(* IEC 61131-3 sources: sis-interlock-demo/tests/POUs/Generated/FB_VoteTruth_Test (part 2) *)

(* ---- Fb2oo2DADIMatchesTable.method.impl.st ---- *)
// AUTO-GENERATED by cemgen 1.0.0 — не редактировать: правьте матрицу и запустите
//   python -m cemgen generate <файл матрицы .csv или .xlsx>
// Матрица: SIS-V101-CEM, объект V-101, ревизия B от 2026-10-19, SHA-256 сетки df2ed4841a9453ca
coUnit.TEST('VoteTruth_Fb2oo2DADI_MatchesTable');
stCfg.eArch := E_VoteArch.Vote2oo2;
stCfg.ePolicy := E_DegradePolicy.DegradeAvailable;
stCfg.eInput := E_SisInputKind.Discrete;
stCfg.xDiHealthy := TRUE;
stCfg.eLimitDir := E_LimitDir.High;
stCfg.rTripLimit_eu := 50.0;
stCfg.rHyst_eu := 0.0;
stCfg.rDiscrepancyMax_eu := 0.0;
stCfg.tDiscrepancyDelay := T#0S;
stCfg.tBypassMax := T#1H;
stCfg.uiMaxBypass := 1;
FOR uiRow := 0 TO 63 DO
    RowInputs(uiRow := uiRow, uiChannels := 2, xBypass := FALSE, stIn := stIn, stCmd := stCmd);
    fbVote(stIn := stIn, stCmd := stCmd, stCfg := stCfg, xBypassPermit := TRUE, uiCause := 1,
        itfTime := fbTime);
    RowInputs(uiRow := uiRow, uiChannels := 2, xBypass := TRUE, stIn := stIn, stCmd := stCmd);
    fbVote(stIn := stIn, stCmd := stCmd, stCfg := stCfg, xBypassPermit := TRUE, uiCause := 1,
        itfTime := fbTime);
    bAct := EncodeFb(xTrip := fbVote.xTrip, stSts := fbVote.stSts);
    bExp := GVL_VoteTruthTable.TT_FB_2OO2_DA_DI[uiRow];
    xMiss := bAct <> bExp;
    xFirst := xMiss AND uiMismatch = 0;
    uiFirstRow := SEL(xFirst, uiFirstRow, uiRow);
    bFirstExp := SEL(xFirst, bFirstExp, bExp);
    bFirstAct := SEL(xFirst, bFirstAct, bAct);
    uiMismatch := uiMismatch + BOOL_TO_UINT(xMiss);
END_FOR
AssertEquals_UINT(Expected := 0, Actual := uiMismatch,
    Message := MismatchText(sTable := 'TT_FB_2OO2_DA_DI', uiRow := uiFirstRow, bExpected := bFirstExp,
        bActual := bFirstAct));
coUnit.TEST_FINISHED();

(* ---- Fb2oo2DSAIMatchesTable.method.decl.st ---- *)
// AUTO-GENERATED by cemgen 1.0.0 — не редактировать: правьте матрицу и запустите
//   python -m cemgen generate <файл матрицы .csv или .xlsx>
// Матрица: SIS-V101-CEM, объект V-101, ревизия B от 2026-10-19, SHA-256 сетки df2ed4841a9453ca
// Назначение: тест VoteTruth_Fb2oo2DSAI_MatchesTable набора FB_VoteTruth_Test.
// Автор:      kr0nsch; код — генератор cemgen
// Версия:     1.0.0
// Документ:   docs/DESIGN.md, раздел «10. Генератор cemgen»; docs/cause_effect_matrix.md
// ВНИМАНИЕ:   код демонстрационный и не предназначен для систем безопасности. Реальная ПАЗ требует
//             определения SIL, сертифицированных аппаратных и программных средств и валидации по
//             ГОСТ Р МЭК 61511.
// FB_Voting, схема 2oo2, политика DegradeSafe, аналоговые каналы: все 64 сочетаний «требование ×
// достоверность × запрос байпаса» совпадают с таблицей TT_FB_2OO2_DS_AI. На строку — два вызова одного
// экземпляра: без запросов байпаса (сброс байпасов прошлой строки) и с полной строкой.
METHOD PRIVATE Fb2oo2DSAIMatchesTable
VAR
    fbTime     : PL.FB_FakeTime;   // время не меняется
    fbVote     : FB_Voting;        // ФБ под тестом, один экземпляр на все строки
    stCfg      : ST_VotingCfg;     // конфигурация теста уровня 2
    stIn       : ST_VoteIn;        // входы строки
    stCmd      : ST_VoteCmd;       // запросы байпаса строки
    uiRow      : UINT;             // строка таблицы
    bAct       : BYTE;             // фактический байт результата
    bExp       : BYTE;             // ожидаемый байт из таблицы
    xMiss      : BOOL;             // строка не совпала
    xFirst     : BOOL;             // первая несовпавшая строка
    uiMismatch : UINT;             // несовпавших строк
    uiFirstRow : UINT;             // первая несовпавшая строка
    bFirstExp  : BYTE;             // ожидаемый байт первой несовпавшей строки
    bFirstAct  : BYTE;             // фактический байт первой несовпавшей строки
END_VAR

(* ---- Fb2oo2DSAIMatchesTable.method.impl.st ---- *)
// AUTO-GENERATED by cemgen 1.0.0 — не редактировать: правьте матрицу и запустите
//   python -m cemgen generate <файл матрицы .csv или .xlsx>
// Матрица: SIS-V101-CEM, объект V-101, ревизия B от 2026-10-19, SHA-256 сетки df2ed4841a9453ca
coUnit.TEST('VoteTruth_Fb2oo2DSAI_MatchesTable');
stCfg.eArch := E_VoteArch.Vote2oo2;
stCfg.ePolicy := E_DegradePolicy.DegradeSafe;
stCfg.eInput := E_SisInputKind.Analog;
stCfg.xDiHealthy := TRUE;
stCfg.eLimitDir := E_LimitDir.High;
stCfg.rTripLimit_eu := 50.0;
stCfg.rHyst_eu := 0.0;
stCfg.rDiscrepancyMax_eu := 0.0;
stCfg.tDiscrepancyDelay := T#0S;
stCfg.tBypassMax := T#1H;
stCfg.uiMaxBypass := 1;
FOR uiRow := 0 TO 63 DO
    RowInputs(uiRow := uiRow, uiChannels := 2, xBypass := FALSE, stIn := stIn, stCmd := stCmd);
    fbVote(stIn := stIn, stCmd := stCmd, stCfg := stCfg, xBypassPermit := TRUE, uiCause := 1,
        itfTime := fbTime);
    RowInputs(uiRow := uiRow, uiChannels := 2, xBypass := TRUE, stIn := stIn, stCmd := stCmd);
    fbVote(stIn := stIn, stCmd := stCmd, stCfg := stCfg, xBypassPermit := TRUE, uiCause := 1,
        itfTime := fbTime);
    bAct := EncodeFb(xTrip := fbVote.xTrip, stSts := fbVote.stSts);
    bExp := GVL_VoteTruthTable.TT_FB_2OO2_DS_AI[uiRow];
    xMiss := bAct <> bExp;
    xFirst := xMiss AND uiMismatch = 0;
    uiFirstRow := SEL(xFirst, uiFirstRow, uiRow);
    bFirstExp := SEL(xFirst, bFirstExp, bExp);
    bFirstAct := SEL(xFirst, bFirstAct, bAct);
    uiMismatch := uiMismatch + BOOL_TO_UINT(xMiss);
END_FOR
AssertEquals_UINT(Expected := 0, Actual := uiMismatch,
    Message := MismatchText(sTable := 'TT_FB_2OO2_DS_AI', uiRow := uiFirstRow, bExpected := bFirstExp,
        bActual := bFirstAct));
coUnit.TEST_FINISHED();

(* ---- Fb2oo2DSDIMatchesTable.method.decl.st ---- *)
// AUTO-GENERATED by cemgen 1.0.0 — не редактировать: правьте матрицу и запустите
//   python -m cemgen generate <файл матрицы .csv или .xlsx>
// Матрица: SIS-V101-CEM, объект V-101, ревизия B от 2026-10-19, SHA-256 сетки df2ed4841a9453ca
// Назначение: тест VoteTruth_Fb2oo2DSDI_MatchesTable набора FB_VoteTruth_Test.
// Автор:      kr0nsch; код — генератор cemgen
// Версия:     1.0.0
// Документ:   docs/DESIGN.md, раздел «10. Генератор cemgen»; docs/cause_effect_matrix.md
// ВНИМАНИЕ:   код демонстрационный и не предназначен для систем безопасности. Реальная ПАЗ требует
//             определения SIL, сертифицированных аппаратных и программных средств и валидации по
//             ГОСТ Р МЭК 61511.
// FB_Voting, схема 2oo2, политика DegradeSafe, дискретные каналы: все 64 сочетаний «требование ×
// достоверность × запрос байпаса» совпадают с таблицей TT_FB_2OO2_DS_DI. На строку — два вызова одного
// экземпляра: без запросов байпаса (сброс байпасов прошлой строки) и с полной строкой.
METHOD PRIVATE Fb2oo2DSDIMatchesTable
VAR
    fbTime     : PL.FB_FakeTime;   // время не меняется
    fbVote     : FB_Voting;        // ФБ под тестом, один экземпляр на все строки
    stCfg      : ST_VotingCfg;     // конфигурация теста уровня 2
    stIn       : ST_VoteIn;        // входы строки
    stCmd      : ST_VoteCmd;       // запросы байпаса строки
    uiRow      : UINT;             // строка таблицы
    bAct       : BYTE;             // фактический байт результата
    bExp       : BYTE;             // ожидаемый байт из таблицы
    xMiss      : BOOL;             // строка не совпала
    xFirst     : BOOL;             // первая несовпавшая строка
    uiMismatch : UINT;             // несовпавших строк
    uiFirstRow : UINT;             // первая несовпавшая строка
    bFirstExp  : BYTE;             // ожидаемый байт первой несовпавшей строки
    bFirstAct  : BYTE;             // фактический байт первой несовпавшей строки
END_VAR

(* ---- Fb2oo2DSDIMatchesTable.method.impl.st ---- *)
// AUTO-GENERATED by cemgen 1.0.0 — не редактировать: правьте матрицу и запустите
//   python -m cemgen generate <файл матрицы .csv или .xlsx>
// Матрица: SIS-V101-CEM, объект V-101, ревизия B от 2026-10-19, SHA-256 сетки df2ed4841a9453ca
coUnit.TEST('VoteTruth_Fb2oo2DSDI_MatchesTable');
stCfg.eArch := E_VoteArch.Vote2oo2;
stCfg.ePolicy := E_DegradePolicy.DegradeSafe;
stCfg.eInput := E_SisInputKind.Discrete;
stCfg.xDiHealthy := TRUE;
stCfg.eLimitDir := E_LimitDir.High;
stCfg.rTripLimit_eu := 50.0;
stCfg.rHyst_eu := 0.0;
stCfg.rDiscrepancyMax_eu := 0.0;
stCfg.tDiscrepancyDelay := T#0S;
stCfg.tBypassMax := T#1H;
stCfg.uiMaxBypass := 1;
FOR uiRow := 0 TO 63 DO
    RowInputs(uiRow := uiRow, uiChannels := 2, xBypass := FALSE, stIn := stIn, stCmd := stCmd);
    fbVote(stIn := stIn, stCmd := stCmd, stCfg := stCfg, xBypassPermit := TRUE, uiCause := 1,
        itfTime := fbTime);
    RowInputs(uiRow := uiRow, uiChannels := 2, xBypass := TRUE, stIn := stIn, stCmd := stCmd);
    fbVote(stIn := stIn, stCmd := stCmd, stCfg := stCfg, xBypassPermit := TRUE, uiCause := 1,
        itfTime := fbTime);
    bAct := EncodeFb(xTrip := fbVote.xTrip, stSts := fbVote.stSts);
    bExp := GVL_VoteTruthTable.TT_FB_2OO2_DS_DI[uiRow];
    xMiss := bAct <> bExp;
    xFirst := xMiss AND uiMismatch = 0;
    uiFirstRow := SEL(xFirst, uiFirstRow, uiRow);
    bFirstExp := SEL(xFirst, bFirstExp, bExp);
    bFirstAct := SEL(xFirst, bFirstAct, bAct);
    uiMismatch := uiMismatch + BOOL_TO_UINT(xMiss);
END_FOR
AssertEquals_UINT(Expected := 0, Actual := uiMismatch,
    Message := MismatchText(sTable := 'TT_FB_2OO2_DS_DI', uiRow := uiFirstRow, bExpected := bFirstExp,
        bActual := bFirstAct));
coUnit.TEST_FINISHED();

(* ---- Fb2oo2VTAIMatchesTable.method.decl.st ---- *)
// AUTO-GENERATED by cemgen 1.0.0 — не редактировать: правьте матрицу и запустите
//   python -m cemgen generate <файл матрицы .csv или .xlsx>
// Матрица: SIS-V101-CEM, объект V-101, ревизия B от 2026-10-19, SHA-256 сетки df2ed4841a9453ca
// Назначение: тест VoteTruth_Fb2oo2VTAI_MatchesTable набора FB_VoteTruth_Test.
// Автор:      kr0nsch; код — генератор cemgen
// Версия:     1.0.0
// Документ:   docs/DESIGN.md, раздел «10. Генератор cemgen»; docs/cause_effect_matrix.md
// ВНИМАНИЕ:   код демонстрационный и не предназначен для систем безопасности. Реальная ПАЗ требует
//             определения SIL, сертифицированных аппаратных и программных средств и валидации по
//             ГОСТ Р МЭК 61511.
// FB_Voting, схема 2oo2, политика VoteTrip, аналоговые каналы: все 64 сочетаний «требование ×
// достоверность × запрос байпаса» совпадают с таблицей TT_FB_2OO2_VT_AI. На строку — два вызова одного
// экземпляра: без запросов байпаса (сброс байпасов прошлой строки) и с полной строкой.
METHOD PRIVATE Fb2oo2VTAIMatchesTable
VAR
    fbTime     : PL.FB_FakeTime;   // время не меняется
    fbVote     : FB_Voting;        // ФБ под тестом, один экземпляр на все строки
    stCfg      : ST_VotingCfg;     // конфигурация теста уровня 2
    stIn       : ST_VoteIn;        // входы строки
    stCmd      : ST_VoteCmd;       // запросы байпаса строки
    uiRow      : UINT;             // строка таблицы
    bAct       : BYTE;             // фактический байт результата
    bExp       : BYTE;             // ожидаемый байт из таблицы
    xMiss      : BOOL;             // строка не совпала
    xFirst     : BOOL;             // первая несовпавшая строка
    uiMismatch : UINT;             // несовпавших строк
    uiFirstRow : UINT;             // первая несовпавшая строка
    bFirstExp  : BYTE;             // ожидаемый байт первой несовпавшей строки
    bFirstAct  : BYTE;             // фактический байт первой несовпавшей строки
END_VAR

(* ---- Fb2oo2VTAIMatchesTable.method.impl.st ---- *)
// AUTO-GENERATED by cemgen 1.0.0 — не редактировать: правьте матрицу и запустите
//   python -m cemgen generate <файл матрицы .csv или .xlsx>
// Матрица: SIS-V101-CEM, объект V-101, ревизия B от 2026-10-19, SHA-256 сетки df2ed4841a9453ca
coUnit.TEST('VoteTruth_Fb2oo2VTAI_MatchesTable');
stCfg.eArch := E_VoteArch.Vote2oo2;
stCfg.ePolicy := E_DegradePolicy.VoteTrip;
stCfg.eInput := E_SisInputKind.Analog;
stCfg.xDiHealthy := TRUE;
stCfg.eLimitDir := E_LimitDir.High;
stCfg.rTripLimit_eu := 50.0;
stCfg.rHyst_eu := 0.0;
stCfg.rDiscrepancyMax_eu := 0.0;
stCfg.tDiscrepancyDelay := T#0S;
stCfg.tBypassMax := T#1H;
stCfg.uiMaxBypass := 1;
FOR uiRow := 0 TO 63 DO
    RowInputs(uiRow := uiRow, uiChannels := 2, xBypass := FALSE, stIn := stIn, stCmd := stCmd);
    fbVote(stIn := stIn, stCmd := stCmd, stCfg := stCfg, xBypassPermit := TRUE, uiCause := 1,
        itfTime := fbTime);
    RowInputs(uiRow := uiRow, uiChannels := 2, xBypass := TRUE, stIn := stIn, stCmd := stCmd);
    fbVote(stIn := stIn, stCmd := stCmd, stCfg := stCfg, xBypassPermit := TRUE, uiCause := 1,
        itfTime := fbTime);
    bAct := EncodeFb(xTrip := fbVote.xTrip, stSts := fbVote.stSts);
    bExp := GVL_VoteTruthTable.TT_FB_2OO2_VT_AI[uiRow];
    xMiss := bAct <> bExp;
    xFirst := xMiss AND uiMismatch = 0;
    uiFirstRow := SEL(xFirst, uiFirstRow, uiRow);
    bFirstExp := SEL(xFirst, bFirstExp, bExp);
    bFirstAct := SEL(xFirst, bFirstAct, bAct);
    uiMismatch := uiMismatch + BOOL_TO_UINT(xMiss);
END_FOR
AssertEquals_UINT(Expected := 0, Actual := uiMismatch,
    Message := MismatchText(sTable := 'TT_FB_2OO2_VT_AI', uiRow := uiFirstRow, bExpected := bFirstExp,
        bActual := bFirstAct));
coUnit.TEST_FINISHED();

(* ---- Fb2oo2VTDIMatchesTable.method.decl.st ---- *)
// AUTO-GENERATED by cemgen 1.0.0 — не редактировать: правьте матрицу и запустите
//   python -m cemgen generate <файл матрицы .csv или .xlsx>
// Матрица: SIS-V101-CEM, объект V-101, ревизия B от 2026-10-19, SHA-256 сетки df2ed4841a9453ca
// Назначение: тест VoteTruth_Fb2oo2VTDI_MatchesTable набора FB_VoteTruth_Test.
// Автор:      kr0nsch; код — генератор cemgen
// Версия:     1.0.0
// Документ:   docs/DESIGN.md, раздел «10. Генератор cemgen»; docs/cause_effect_matrix.md
// ВНИМАНИЕ:   код демонстрационный и не предназначен для систем безопасности. Реальная ПАЗ требует
//             определения SIL, сертифицированных аппаратных и программных средств и валидации по
//             ГОСТ Р МЭК 61511.
// FB_Voting, схема 2oo2, политика VoteTrip, дискретные каналы: все 64 сочетаний «требование ×
// достоверность × запрос байпаса» совпадают с таблицей TT_FB_2OO2_VT_DI. На строку — два вызова одного
// экземпляра: без запросов байпаса (сброс байпасов прошлой строки) и с полной строкой.
METHOD PRIVATE Fb2oo2VTDIMatchesTable
VAR
    fbTime     : PL.FB_FakeTime;   // время не меняется
    fbVote     : FB_Voting;        // ФБ под тестом, один экземпляр на все строки
    stCfg      : ST_VotingCfg;     // конфигурация теста уровня 2
    stIn       : ST_VoteIn;        // входы строки
    stCmd      : ST_VoteCmd;       // запросы байпаса строки
    uiRow      : UINT;             // строка таблицы
    bAct       : BYTE;             // фактический байт результата
    bExp       : BYTE;             // ожидаемый байт из таблицы
    xMiss      : BOOL;             // строка не совпала
    xFirst     : BOOL;             // первая несовпавшая строка
    uiMismatch : UINT;             // несовпавших строк
    uiFirstRow : UINT;             // первая несовпавшая строка
    bFirstExp  : BYTE;             // ожидаемый байт первой несовпавшей строки
    bFirstAct  : BYTE;             // фактический байт первой несовпавшей строки
END_VAR

(* ---- Fb2oo2VTDIMatchesTable.method.impl.st ---- *)
// AUTO-GENERATED by cemgen 1.0.0 — не редактировать: правьте матрицу и запустите
//   python -m cemgen generate <файл матрицы .csv или .xlsx>
// Матрица: SIS-V101-CEM, объект V-101, ревизия B от 2026-10-19, SHA-256 сетки df2ed4841a9453ca
coUnit.TEST('VoteTruth_Fb2oo2VTDI_MatchesTable');
stCfg.eArch := E_VoteArch.Vote2oo2;
stCfg.ePolicy := E_DegradePolicy.VoteTrip;
stCfg.eInput := E_SisInputKind.Discrete;
stCfg.xDiHealthy := TRUE;
stCfg.eLimitDir := E_LimitDir.High;
stCfg.rTripLimit_eu := 50.0;
stCfg.rHyst_eu := 0.0;
stCfg.rDiscrepancyMax_eu := 0.0;
stCfg.tDiscrepancyDelay := T#0S;
stCfg.tBypassMax := T#1H;
stCfg.uiMaxBypass := 1;
FOR uiRow := 0 TO 63 DO
    RowInputs(uiRow := uiRow, uiChannels := 2, xBypass := FALSE, stIn := stIn, stCmd := stCmd);
    fbVote(stIn := stIn, stCmd := stCmd, stCfg := stCfg, xBypassPermit := TRUE, uiCause := 1,
        itfTime := fbTime);
    RowInputs(uiRow := uiRow, uiChannels := 2, xBypass := TRUE, stIn := stIn, stCmd := stCmd);
    fbVote(stIn := stIn, stCmd := stCmd, stCfg := stCfg, xBypassPermit := TRUE, uiCause := 1,
        itfTime := fbTime);
    bAct := EncodeFb(xTrip := fbVote.xTrip, stSts := fbVote.stSts);
    bExp := GVL_VoteTruthTable.TT_FB_2OO2_VT_DI[uiRow];
    xMiss := bAct <> bExp;
    xFirst := xMiss AND uiMismatch = 0;
    uiFirstRow := SEL(xFirst, uiFirstRow, uiRow);
    bFirstExp := SEL(xFirst, bFirstExp, bExp);
    bFirstAct := SEL(xFirst, bFirstAct, bAct);
    uiMismatch := uiMismatch + BOOL_TO_UINT(xMiss);
END_FOR
AssertEquals_UINT(Expected := 0, Actual := uiMismatch,
    Message := MismatchText(sTable := 'TT_FB_2OO2_VT_DI', uiRow := uiFirstRow, bExpected := bFirstExp,
        bActual := bFirstAct));
coUnit.TEST_FINISHED();

(* ---- Fb2oo3DAAIMatchesTable.method.decl.st ---- *)
// AUTO-GENERATED by cemgen 1.0.0 — не редактировать: правьте матрицу и запустите
//   python -m cemgen generate <файл матрицы .csv или .xlsx>
// Матрица: SIS-V101-CEM, объект V-101, ревизия B от 2026-10-19, SHA-256 сетки df2ed4841a9453ca
// Назначение: тест VoteTruth_Fb2oo3DAAI_MatchesTable набора FB_VoteTruth_Test.
// Автор:      kr0nsch; код — генератор cemgen
// Версия:     1.0.0
// Документ:   docs/DESIGN.md, раздел «10. Генератор cemgen»; docs/cause_effect_matrix.md
// ВНИМАНИЕ:   код демонстрационный и не предназначен для систем безопасности. Реальная ПАЗ требует
//             определения SIL, сертифицированных аппаратных и программных средств и валидации по
//             ГОСТ Р МЭК 61511.
// FB_Voting, схема 2oo3, политика DegradeAvailable, аналоговые каналы: все 512 сочетаний «требование ×
// достоверность × запрос байпаса» совпадают с таблицей TT_FB_2OO3_DA_AI. На строку — два вызова одного
// экземпляра: без запросов байпаса (сброс байпасов прошлой строки) и с полной строкой.
METHOD PRIVATE Fb2oo3DAAIMatchesTable
VAR
    fbTime     : PL.FB_FakeTime;   // время не меняется
    fbVote     : FB_Voting;        // ФБ под тестом, один экземпляр на все строки
    stCfg      : ST_VotingCfg;     // конфигурация теста уровня 2
    stIn       : ST_VoteIn;        // входы строки
    stCmd      : ST_VoteCmd;       // запросы байпаса строки
    uiRow      : UINT;             // строка таблицы
    bAct       : BYTE;             // фактический байт результата
    bExp       : BYTE;             // ожидаемый байт из таблицы
    xMiss      : BOOL;             // строка не совпала
    xFirst     : BOOL;             // первая несовпавшая строка
    uiMismatch : UINT;             // несовпавших строк
    uiFirstRow : UINT;             // первая несовпавшая строка
    bFirstExp  : BYTE;             // ожидаемый байт первой несовпавшей строки
    bFirstAct  : BYTE;             // фактический байт первой несовпавшей строки
END_VAR

(* ---- Fb2oo3DAAIMatchesTable.method.impl.st ---- *)
// AUTO-GENERATED by cemgen 1.0.0 — не редактировать: правьте матрицу и запустите
//   python -m cemgen generate <файл матрицы .csv или .xlsx>
// Матрица: SIS-V101-CEM, объект V-101, ревизия B от 2026-10-19, SHA-256 сетки df2ed4841a9453ca
coUnit.TEST('VoteTruth_Fb2oo3DAAI_MatchesTable');
stCfg.eArch := E_VoteArch.Vote2oo3;
stCfg.ePolicy := E_DegradePolicy.DegradeAvailable;
stCfg.eInput := E_SisInputKind.Analog;
stCfg.xDiHealthy := TRUE;
stCfg.eLimitDir := E_LimitDir.High;
stCfg.rTripLimit_eu := 50.0;
stCfg.rHyst_eu := 0.0;
stCfg.rDiscrepancyMax_eu := 0.0;
stCfg.tDiscrepancyDelay := T#0S;
stCfg.tBypassMax := T#1H;
stCfg.uiMaxBypass := 1;
FOR uiRow := 0 TO 511 DO
    RowInputs(uiRow := uiRow, uiChannels := 3, xBypass := FALSE, stIn := stIn, stCmd := stCmd);
    fbVote(stIn := stIn, stCmd := stCmd, stCfg := stCfg, xBypassPermit := TRUE, uiCause := 1,
        itfTime := fbTime);
    RowInputs(uiRow := uiRow, uiChannels := 3, xBypass := TRUE, stIn := stIn, stCmd := stCmd);
    fbVote(stIn := stIn, stCmd := stCmd, stCfg := stCfg, xBypassPermit := TRUE, uiCause := 1,
        itfTime := fbTime);
    bAct := EncodeFb(xTrip := fbVote.xTrip, stSts := fbVote.stSts);
    bExp := GVL_VoteTruthTable.TT_FB_2OO3_DA_AI[uiRow];
    xMiss := bAct <> bExp;
    xFirst := xMiss AND uiMismatch = 0;
    uiFirstRow := SEL(xFirst, uiFirstRow, uiRow);
    bFirstExp := SEL(xFirst, bFirstExp, bExp);
    bFirstAct := SEL(xFirst, bFirstAct, bAct);
    uiMismatch := uiMismatch + BOOL_TO_UINT(xMiss);
END_FOR
AssertEquals_UINT(Expected := 0, Actual := uiMismatch,
    Message := MismatchText(sTable := 'TT_FB_2OO3_DA_AI', uiRow := uiFirstRow, bExpected := bFirstExp,
        bActual := bFirstAct));
coUnit.TEST_FINISHED();

(* ---- Fb2oo3DADIMatchesTable.method.decl.st ---- *)
// AUTO-GENERATED by cemgen 1.0.0 — не редактировать: правьте матрицу и запустите
//   python -m cemgen generate <файл матрицы .csv или .xlsx>
// Матрица: SIS-V101-CEM, объект V-101, ревизия B от 2026-10-19, SHA-256 сетки df2ed4841a9453ca
// Назначение: тест VoteTruth_Fb2oo3DADI_MatchesTable набора FB_VoteTruth_Test.
// Автор:      kr0nsch; код — генератор cemgen
// Версия:     1.0.0
// Документ:   docs/DESIGN.md, раздел «10. Генератор cemgen»; docs/cause_effect_matrix.md
// ВНИМАНИЕ:   код демонстрационный и не предназначен для систем безопасности. Реальная ПАЗ требует
//             определения SIL, сертифицированных аппаратных и программных средств и валидации по
//             ГОСТ Р МЭК 61511.
// FB_Voting, схема 2oo3, политика DegradeAvailable, дискретные каналы: все 512 сочетаний «требование ×
// достоверность × запрос байпаса» совпадают с таблицей TT_FB_2OO3_DA_DI. На строку — два вызова одного
// экземпляра: без запросов байпаса (сброс байпасов прошлой строки) и с полной строкой.
METHOD PRIVATE Fb2oo3DADIMatchesTable
VAR
    fbTime     : PL.FB_FakeTime;   // время не меняется
    fbVote     : FB_Voting;        // ФБ под тестом, один экземпляр на все строки
    stCfg      : ST_VotingCfg;     // конфигурация теста уровня 2
    stIn       : ST_VoteIn;        // входы строки
    stCmd      : ST_VoteCmd;       // запросы байпаса строки
    uiRow      : UINT;             // строка таблицы
    bAct       : BYTE;             // фактический байт результата
    bExp       : BYTE;             // ожидаемый байт из таблицы
    xMiss      : BOOL;             // строка не совпала
    xFirst     : BOOL;             // первая несовпавшая строка
    uiMismatch : UINT;             // несовпавших строк
    uiFirstRow : UINT;             // первая несовпавшая строка
    bFirstExp  : BYTE;             // ожидаемый байт первой несовпавшей строки
    bFirstAct  : BYTE;             // фактический байт первой несовпавшей строки
END_VAR

(* ---- Fb2oo3DADIMatchesTable.method.impl.st ---- *)
// AUTO-GENERATED by cemgen 1.0.0 — не редактировать: правьте матрицу и запустите
//   python -m cemgen generate <файл матрицы .csv или .xlsx>
// Матрица: SIS-V101-CEM, объект V-101, ревизия B от 2026-10-19, SHA-256 сетки df2ed4841a9453ca
coUnit.TEST('VoteTruth_Fb2oo3DADI_MatchesTable');
stCfg.eArch := E_VoteArch.Vote2oo3;
stCfg.ePolicy := E_DegradePolicy.DegradeAvailable;
stCfg.eInput := E_SisInputKind.Discrete;
stCfg.xDiHealthy := TRUE;
stCfg.eLimitDir := E_LimitDir.High;
stCfg.rTripLimit_eu := 50.0;
stCfg.rHyst_eu := 0.0;
stCfg.rDiscrepancyMax_eu := 0.0;
stCfg.tDiscrepancyDelay := T#0S;
stCfg.tBypassMax := T#1H;
stCfg.uiMaxBypass := 1;
FOR uiRow := 0 TO 511 DO
    RowInputs(uiRow := uiRow, uiChannels := 3, xBypass := FALSE, stIn := stIn, stCmd := stCmd);
    fbVote(stIn := stIn, stCmd := stCmd, stCfg := stCfg, xBypassPermit := TRUE, uiCause := 1,
        itfTime := fbTime);
    RowInputs(uiRow := uiRow, uiChannels := 3, xBypass := TRUE, stIn := stIn, stCmd := stCmd);
    fbVote(stIn := stIn, stCmd := stCmd, stCfg := stCfg, xBypassPermit := TRUE, uiCause := 1,
        itfTime := fbTime);
    bAct := EncodeFb(xTrip := fbVote.xTrip, stSts := fbVote.stSts);
    bExp := GVL_VoteTruthTable.TT_FB_2OO3_DA_DI[uiRow];
    xMiss := bAct <> bExp;
    xFirst := xMiss AND uiMismatch = 0;
    uiFirstRow := SEL(xFirst, uiFirstRow, uiRow);
    bFirstExp := SEL(xFirst, bFirstExp, bExp);
    bFirstAct := SEL(xFirst, bFirstAct, bAct);
    uiMismatch := uiMismatch + BOOL_TO_UINT(xMiss);
END_FOR
AssertEquals_UINT(Expected := 0, Actual := uiMismatch,
    Message := MismatchText(sTable := 'TT_FB_2OO3_DA_DI', uiRow := uiFirstRow, bExpected := bFirstExp,
        bActual := bFirstAct));
coUnit.TEST_FINISHED();

(* ---- Fb2oo3DSAIMatchesTable.method.decl.st ---- *)
// AUTO-GENERATED by cemgen 1.0.0 — не редактировать: правьте матрицу и запустите
//   python -m cemgen generate <файл матрицы .csv или .xlsx>
// Матрица: SIS-V101-CEM, объект V-101, ревизия B от 2026-10-19, SHA-256 сетки df2ed4841a9453ca
// Назначение: тест VoteTruth_Fb2oo3DSAI_MatchesTable набора FB_VoteTruth_Test.
// Автор:      kr0nsch; код — генератор cemgen
// Версия:     1.0.0
// Документ:   docs/DESIGN.md, раздел «10. Генератор cemgen»; docs/cause_effect_matrix.md
// ВНИМАНИЕ:   код демонстрационный и не предназначен для систем безопасности. Реальная ПАЗ требует
//             определения SIL, сертифицированных аппаратных и программных средств и валидации по
//             ГОСТ Р МЭК 61511.
// FB_Voting, схема 2oo3, политика DegradeSafe, аналоговые каналы: все 512 сочетаний «требование ×
// достоверность × запрос байпаса» совпадают с таблицей TT_FB_2OO3_DS_AI. На строку — два вызова одного
// экземпляра: без запросов байпаса (сброс байпасов прошлой строки) и с полной строкой.
METHOD PRIVATE Fb2oo3DSAIMatchesTable
VAR
    fbTime     : PL.FB_FakeTime;   // время не меняется
    fbVote     : FB_Voting;        // ФБ под тестом, один экземпляр на все строки
    stCfg      : ST_VotingCfg;     // конфигурация теста уровня 2
    stIn       : ST_VoteIn;        // входы строки
    stCmd      : ST_VoteCmd;       // запросы байпаса строки
    uiRow      : UINT;             // строка таблицы
    bAct       : BYTE;             // фактический байт результата
    bExp       : BYTE;             // ожидаемый байт из таблицы
    xMiss      : BOOL;             // строка не совпала
    xFirst     : BOOL;             // первая несовпавшая строка
    uiMismatch : UINT;             // несовпавших строк
    uiFirstRow : UINT;             // первая несовпавшая строка
    bFirstExp  : BYTE;             // ожидаемый байт первой несовпавшей строки
    bFirstAct  : BYTE;             // фактический байт первой несовпавшей строки
END_VAR

(* ---- Fb2oo3DSAIMatchesTable.method.impl.st ---- *)
// AUTO-GENERATED by cemgen 1.0.0 — не редактировать: правьте матрицу и запустите
//   python -m cemgen generate <файл матрицы .csv или .xlsx>
// Матрица: SIS-V101-CEM, объект V-101, ревизия B от 2026-10-19, SHA-256 сетки df2ed4841a9453ca
coUnit.TEST('VoteTruth_Fb2oo3DSAI_MatchesTable');
stCfg.eArch := E_VoteArch.Vote2oo3;
stCfg.ePolicy := E_DegradePolicy.DegradeSafe;
stCfg.eInput := E_SisInputKind.Analog;
stCfg.xDiHealthy := TRUE;
stCfg.eLimitDir := E_LimitDir.High;
stCfg.rTripLimit_eu := 50.0;
stCfg.rHyst_eu := 0.0;
stCfg.rDiscrepancyMax_eu := 0.0;
stCfg.tDiscrepancyDelay := T#0S;
stCfg.tBypassMax := T#1H;
stCfg.uiMaxBypass := 1;
FOR uiRow := 0 TO 511 DO
    RowInputs(uiRow := uiRow, uiChannels := 3, xBypass := FALSE, stIn := stIn, stCmd := stCmd);
    fbVote(stIn := stIn, stCmd := stCmd, stCfg := stCfg, xBypassPermit := TRUE, uiCause := 1,
        itfTime := fbTime);
    RowInputs(uiRow := uiRow, uiChannels := 3, xBypass := TRUE, stIn := stIn, stCmd := stCmd);
    fbVote(stIn := stIn, stCmd := stCmd, stCfg := stCfg, xBypassPermit := TRUE, uiCause := 1,
        itfTime := fbTime);
    bAct := EncodeFb(xTrip := fbVote.xTrip, stSts := fbVote.stSts);
    bExp := GVL_VoteTruthTable.TT_FB_2OO3_DS_AI[uiRow];
    xMiss := bAct <> bExp;
    xFirst := xMiss AND uiMismatch = 0;
    uiFirstRow := SEL(xFirst, uiFirstRow, uiRow);
    bFirstExp := SEL(xFirst, bFirstExp, bExp);
    bFirstAct := SEL(xFirst, bFirstAct, bAct);
    uiMismatch := uiMismatch + BOOL_TO_UINT(xMiss);
END_FOR
AssertEquals_UINT(Expected := 0, Actual := uiMismatch,
    Message := MismatchText(sTable := 'TT_FB_2OO3_DS_AI', uiRow := uiFirstRow, bExpected := bFirstExp,
        bActual := bFirstAct));
coUnit.TEST_FINISHED();

(* ---- Fb2oo3DSDIMatchesTable.method.decl.st ---- *)
// AUTO-GENERATED by cemgen 1.0.0 — не редактировать: правьте матрицу и запустите
//   python -m cemgen generate <файл матрицы .csv или .xlsx>
// Матрица: SIS-V101-CEM, объект V-101, ревизия B от 2026-10-19, SHA-256 сетки df2ed4841a9453ca
// Назначение: тест VoteTruth_Fb2oo3DSDI_MatchesTable набора FB_VoteTruth_Test.
// Автор:      kr0nsch; код — генератор cemgen
// Версия:     1.0.0
// Документ:   docs/DESIGN.md, раздел «10. Генератор cemgen»; docs/cause_effect_matrix.md
// ВНИМАНИЕ:   код демонстрационный и не предназначен для систем безопасности. Реальная ПАЗ требует
//             определения SIL, сертифицированных аппаратных и программных средств и валидации по
//             ГОСТ Р МЭК 61511.
// FB_Voting, схема 2oo3, политика DegradeSafe, дискретные каналы: все 512 сочетаний «требование ×
// достоверность × запрос байпаса» совпадают с таблицей TT_FB_2OO3_DS_DI. На строку — два вызова одного
// экземпляра: без запросов байпаса (сброс байпасов прошлой строки) и с полной строкой.
METHOD PRIVATE Fb2oo3DSDIMatchesTable
VAR
    fbTime     : PL.FB_FakeTime;   // время не меняется
    fbVote     : FB_Voting;        // ФБ под тестом, один экземпляр на все строки
    stCfg      : ST_VotingCfg;     // конфигурация теста уровня 2
    stIn       : ST_VoteIn;        // входы строки
    stCmd      : ST_VoteCmd;       // запросы байпаса строки
    uiRow      : UINT;             // строка таблицы
    bAct       : BYTE;             // фактический байт результата
    bExp       : BYTE;             // ожидаемый байт из таблицы
    xMiss      : BOOL;             // строка не совпала
    xFirst     : BOOL;             // первая несовпавшая строка
    uiMismatch : UINT;             // несовпавших строк
    uiFirstRow : UINT;             // первая несовпавшая строка
    bFirstExp  : BYTE;             // ожидаемый байт первой несовпавшей строки
    bFirstAct  : BYTE;             // фактический байт первой несовпавшей строки
END_VAR

(* ---- Fb2oo3DSDIMatchesTable.method.impl.st ---- *)
// AUTO-GENERATED by cemgen 1.0.0 — не редактировать: правьте матрицу и запустите
//   python -m cemgen generate <файл матрицы .csv или .xlsx>
// Матрица: SIS-V101-CEM, объект V-101, ревизия B от 2026-10-19, SHA-256 сетки df2ed4841a9453ca
coUnit.TEST('VoteTruth_Fb2oo3DSDI_MatchesTable');
stCfg.eArch := E_VoteArch.Vote2oo3;
stCfg.ePolicy := E_DegradePolicy.DegradeSafe;
stCfg.eInput := E_SisInputKind.Discrete;
stCfg.xDiHealthy := TRUE;
stCfg.eLimitDir := E_LimitDir.High;
stCfg.rTripLimit_eu := 50.0;
stCfg.rHyst_eu := 0.0;
stCfg.rDiscrepancyMax_eu := 0.0;
stCfg.tDiscrepancyDelay := T#0S;
stCfg.tBypassMax := T#1H;
stCfg.uiMaxBypass := 1;
FOR uiRow := 0 TO 511 DO
    RowInputs(uiRow := uiRow, uiChannels := 3, xBypass := FALSE, stIn := stIn, stCmd := stCmd);
    fbVote(stIn := stIn, stCmd := stCmd, stCfg := stCfg, xBypassPermit := TRUE, uiCause := 1,
        itfTime := fbTime);
    RowInputs(uiRow := uiRow, uiChannels := 3, xBypass := TRUE, stIn := stIn, stCmd := stCmd);
    fbVote(stIn := stIn, stCmd := stCmd, stCfg := stCfg, xBypassPermit := TRUE, uiCause := 1,
        itfTime := fbTime);
    bAct := EncodeFb(xTrip := fbVote.xTrip, stSts := fbVote.stSts);
    bExp := GVL_VoteTruthTable.TT_FB_2OO3_DS_DI[uiRow];
    xMiss := bAct <> bExp;
    xFirst := xMiss AND uiMismatch = 0;
    uiFirstRow := SEL(xFirst, uiFirstRow, uiRow);
    bFirstExp := SEL(xFirst, bFirstExp, bExp);
    bFirstAct := SEL(xFirst, bFirstAct, bAct);
    uiMismatch := uiMismatch + BOOL_TO_UINT(xMiss);
END_FOR
AssertEquals_UINT(Expected := 0, Actual := uiMismatch,
    Message := MismatchText(sTable := 'TT_FB_2OO3_DS_DI', uiRow := uiFirstRow, bExpected := bFirstExp,
        bActual := bFirstAct));
coUnit.TEST_FINISHED();

(* ---- Fb2oo3VTAIMatchesTable.method.decl.st ---- *)
// AUTO-GENERATED by cemgen 1.0.0 — не редактировать: правьте матрицу и запустите
//   python -m cemgen generate <файл матрицы .csv или .xlsx>
// Матрица: SIS-V101-CEM, объект V-101, ревизия B от 2026-10-19, SHA-256 сетки df2ed4841a9453ca
// Назначение: тест VoteTruth_Fb2oo3VTAI_MatchesTable набора FB_VoteTruth_Test.
// Автор:      kr0nsch; код — генератор cemgen
// Версия:     1.0.0
// Документ:   docs/DESIGN.md, раздел «10. Генератор cemgen»; docs/cause_effect_matrix.md
// ВНИМАНИЕ:   код демонстрационный и не предназначен для систем безопасности. Реальная ПАЗ требует
//             определения SIL, сертифицированных аппаратных и программных средств и валидации по
//             ГОСТ Р МЭК 61511.
// FB_Voting, схема 2oo3, политика VoteTrip, аналоговые каналы: все 512 сочетаний «требование ×
// достоверность × запрос байпаса» совпадают с таблицей TT_FB_2OO3_VT_AI. На строку — два вызова одного
// экземпляра: без запросов байпаса (сброс байпасов прошлой строки) и с полной строкой.
METHOD PRIVATE Fb2oo3VTAIMatchesTable
VAR
    fbTime     : PL.FB_FakeTime;   // время не меняется
    fbVote     : FB_Voting;        // ФБ под тестом, один экземпляр на все строки
    stCfg      : ST_VotingCfg;     // конфигурация теста уровня 2
    stIn       : ST_VoteIn;        // входы строки
    stCmd      : ST_VoteCmd;       // запросы байпаса строки
    uiRow      : UINT;             // строка таблицы
    bAct       : BYTE;             // фактический байт результата
    bExp       : BYTE;             // ожидаемый байт из таблицы
    xMiss      : BOOL;             // строка не совпала
    xFirst     : BOOL;             // первая несовпавшая строка
    uiMismatch : UINT;             // несовпавших строк
    uiFirstRow : UINT;             // первая несовпавшая строка
    bFirstExp  : BYTE;             // ожидаемый байт первой несовпавшей строки
    bFirstAct  : BYTE;             // фактический байт первой несовпавшей строки
END_VAR

(* ---- Fb2oo3VTAIMatchesTable.method.impl.st ---- *)
// AUTO-GENERATED by cemgen 1.0.0 — не редактировать: правьте матрицу и запустите
//   python -m cemgen generate <файл матрицы .csv или .xlsx>
// Матрица: SIS-V101-CEM, объект V-101, ревизия B от 2026-10-19, SHA-256 сетки df2ed4841a9453ca
coUnit.TEST('VoteTruth_Fb2oo3VTAI_MatchesTable');
stCfg.eArch := E_VoteArch.Vote2oo3;
stCfg.ePolicy := E_DegradePolicy.VoteTrip;
stCfg.eInput := E_SisInputKind.Analog;
stCfg.xDiHealthy := TRUE;
stCfg.eLimitDir := E_LimitDir.High;
stCfg.rTripLimit_eu := 50.0;
stCfg.rHyst_eu := 0.0;
stCfg.rDiscrepancyMax_eu := 0.0;
stCfg.tDiscrepancyDelay := T#0S;
stCfg.tBypassMax := T#1H;
stCfg.uiMaxBypass := 1;
FOR uiRow := 0 TO 511 DO
    RowInputs(uiRow := uiRow, uiChannels := 3, xBypass := FALSE, stIn := stIn, stCmd := stCmd);
    fbVote(stIn := stIn, stCmd := stCmd, stCfg := stCfg, xBypassPermit := TRUE, uiCause := 1,
        itfTime := fbTime);
    RowInputs(uiRow := uiRow, uiChannels := 3, xBypass := TRUE, stIn := stIn, stCmd := stCmd);
    fbVote(stIn := stIn, stCmd := stCmd, stCfg := stCfg, xBypassPermit := TRUE, uiCause := 1,
        itfTime := fbTime);
    bAct := EncodeFb(xTrip := fbVote.xTrip, stSts := fbVote.stSts);
    bExp := GVL_VoteTruthTable.TT_FB_2OO3_VT_AI[uiRow];
    xMiss := bAct <> bExp;
    xFirst := xMiss AND uiMismatch = 0;
    uiFirstRow := SEL(xFirst, uiFirstRow, uiRow);
    bFirstExp := SEL(xFirst, bFirstExp, bExp);
    bFirstAct := SEL(xFirst, bFirstAct, bAct);
    uiMismatch := uiMismatch + BOOL_TO_UINT(xMiss);
END_FOR
AssertEquals_UINT(Expected := 0, Actual := uiMismatch,
    Message := MismatchText(sTable := 'TT_FB_2OO3_VT_AI', uiRow := uiFirstRow, bExpected := bFirstExp,
        bActual := bFirstAct));
coUnit.TEST_FINISHED();

(* ---- Fb2oo3VTDIMatchesTable.method.decl.st ---- *)
// AUTO-GENERATED by cemgen 1.0.0 — не редактировать: правьте матрицу и запустите
//   python -m cemgen generate <файл матрицы .csv или .xlsx>
// Матрица: SIS-V101-CEM, объект V-101, ревизия B от 2026-10-19, SHA-256 сетки df2ed4841a9453ca
// Назначение: тест VoteTruth_Fb2oo3VTDI_MatchesTable набора FB_VoteTruth_Test.
// Автор:      kr0nsch; код — генератор cemgen
// Версия:     1.0.0
// Документ:   docs/DESIGN.md, раздел «10. Генератор cemgen»; docs/cause_effect_matrix.md
// ВНИМАНИЕ:   код демонстрационный и не предназначен для систем безопасности. Реальная ПАЗ требует
//             определения SIL, сертифицированных аппаратных и программных средств и валидации по
//             ГОСТ Р МЭК 61511.
// FB_Voting, схема 2oo3, политика VoteTrip, дискретные каналы: все 512 сочетаний «требование ×
// достоверность × запрос байпаса» совпадают с таблицей TT_FB_2OO3_VT_DI. На строку — два вызова одного
// экземпляра: без запросов байпаса (сброс байпасов прошлой строки) и с полной строкой.
METHOD PRIVATE Fb2oo3VTDIMatchesTable
VAR
    fbTime     : PL.FB_FakeTime;   // время не меняется
    fbVote     : FB_Voting;        // ФБ под тестом, один экземпляр на все строки
    stCfg      : ST_VotingCfg;     // конфигурация теста уровня 2
    stIn       : ST_VoteIn;        // входы строки
    stCmd      : ST_VoteCmd;       // запросы байпаса строки
    uiRow      : UINT;             // строка таблицы
    bAct       : BYTE;             // фактический байт результата
    bExp       : BYTE;             // ожидаемый байт из таблицы
    xMiss      : BOOL;             // строка не совпала
    xFirst     : BOOL;             // первая несовпавшая строка
    uiMismatch : UINT;             // несовпавших строк
    uiFirstRow : UINT;             // первая несовпавшая строка
    bFirstExp  : BYTE;             // ожидаемый байт первой несовпавшей строки
    bFirstAct  : BYTE;             // фактический байт первой несовпавшей строки
END_VAR

(* ---- Fb2oo3VTDIMatchesTable.method.impl.st ---- *)
// AUTO-GENERATED by cemgen 1.0.0 — не редактировать: правьте матрицу и запустите
//   python -m cemgen generate <файл матрицы .csv или .xlsx>
// Матрица: SIS-V101-CEM, объект V-101, ревизия B от 2026-10-19, SHA-256 сетки df2ed4841a9453ca
coUnit.TEST('VoteTruth_Fb2oo3VTDI_MatchesTable');
stCfg.eArch := E_VoteArch.Vote2oo3;
stCfg.ePolicy := E_DegradePolicy.VoteTrip;
stCfg.eInput := E_SisInputKind.Discrete;
stCfg.xDiHealthy := TRUE;
stCfg.eLimitDir := E_LimitDir.High;
stCfg.rTripLimit_eu := 50.0;
stCfg.rHyst_eu := 0.0;
stCfg.rDiscrepancyMax_eu := 0.0;
stCfg.tDiscrepancyDelay := T#0S;
stCfg.tBypassMax := T#1H;
stCfg.uiMaxBypass := 1;
FOR uiRow := 0 TO 511 DO
    RowInputs(uiRow := uiRow, uiChannels := 3, xBypass := FALSE, stIn := stIn, stCmd := stCmd);
    fbVote(stIn := stIn, stCmd := stCmd, stCfg := stCfg, xBypassPermit := TRUE, uiCause := 1,
        itfTime := fbTime);
    RowInputs(uiRow := uiRow, uiChannels := 3, xBypass := TRUE, stIn := stIn, stCmd := stCmd);
    fbVote(stIn := stIn, stCmd := stCmd, stCfg := stCfg, xBypassPermit := TRUE, uiCause := 1,
        itfTime := fbTime);
    bAct := EncodeFb(xTrip := fbVote.xTrip, stSts := fbVote.stSts);
    bExp := GVL_VoteTruthTable.TT_FB_2OO3_VT_DI[uiRow];
    xMiss := bAct <> bExp;
    xFirst := xMiss AND uiMismatch = 0;
    uiFirstRow := SEL(xFirst, uiFirstRow, uiRow);
    bFirstExp := SEL(xFirst, bFirstExp, bExp);
    bFirstAct := SEL(xFirst, bFirstAct, bAct);
    uiMismatch := uiMismatch + BOOL_TO_UINT(xMiss);
END_FOR
AssertEquals_UINT(Expected := 0, Actual := uiMismatch,
    Message := MismatchText(sTable := 'TT_FB_2OO3_VT_DI', uiRow := uiFirstRow, bExpected := bFirstExp,
        bActual := bFirstAct));
coUnit.TEST_FINISHED();

(* ---- MismatchText.method.decl.st ---- *)
// AUTO-GENERATED by cemgen 1.0.0 — не редактировать: правьте матрицу и запустите
//   python -m cemgen generate <файл матрицы .csv или .xlsx>
// Матрица: SIS-V101-CEM, объект V-101, ревизия B от 2026-10-19, SHA-256 сетки df2ed4841a9453ca
// Назначение: вспомогательный метод набора FB_VoteTruth_Test.
// Автор:      kr0nsch; код — генератор cemgen
// Версия:     1.0.0
// Документ:   docs/DESIGN.md, раздел «10. Генератор cemgen»; docs/cause_effect_matrix.md
// ВНИМАНИЕ:   код демонстрационный и не предназначен для систем безопасности. Реальная ПАЗ требует
//             определения SIL, сертифицированных аппаратных и программных средств и валидации по
//             ГОСТ Р МЭК 61511.
// Сообщение ассерта: таблица, первая несовпавшая строка, ожидаемый и фактический байты (ASCII).
METHOD PRIVATE MismatchText : STRING(255)
VAR_INPUT
    sTable    : STRING(40);   // имя таблицы
    uiRow     : UINT;         // первая несовпавшая строка
    bExpected : BYTE;         // ожидаемый байт
    bActual   : BYTE;         // фактический байт
END_VAR
VAR
    sRow      : STRING(12);   // номер строки текстом
    sExpected : STRING(12);   // ожидаемый байт текстом
    sActual   : STRING(12);   // фактический байт текстом
END_VAR

(* ---- RowInputs.method.decl.st ---- *)
// AUTO-GENERATED by cemgen 1.0.0 — не редактировать: правьте матрицу и запустите
//   python -m cemgen generate <файл матрицы .csv или .xlsx>
// Матрица: SIS-V101-CEM, объект V-101, ревизия B от 2026-10-19, SHA-256 сетки df2ed4841a9453ca
// Назначение: вспомогательный метод набора FB_VoteTruth_Test.
// Автор:      kr0nsch; код — генератор cemgen
// Версия:     1.0.0
// Документ:   docs/DESIGN.md, раздел «10. Генератор cemgen»; docs/cause_effect_matrix.md
// ВНИМАНИЕ:   код демонстрационный и не предназначен для систем безопасности. Реальная ПАЗ требует
//             определения SIL, сертифицированных аппаратных и программных средств и валидации по
//             ГОСТ Р МЭК 61511.
// Входы строки уровня 2: для канала k биты 3(k − 1) — требование (DI: axDi := FALSE, AI: 60.0 вместо
// 40.0 при уставке 50.0), +1 — достоверность, +2 — запрос байпаса (только при xBypass). Каналы k > N —
// без требования, недостоверны, без запроса.
METHOD PRIVATE RowInputs
VAR_INPUT
    uiRow      : UINT;   // строка таблицы
    uiChannels : UINT;   // N схемы
    xBypass    : BOOL;   // FALSE — запросы байпаса сняты (первый вызов строки)
END_VAR
VAR_IN_OUT
    stIn  : ST_VoteIn;   // входы группы
    stCmd : ST_VoteCmd;  // запросы байпаса
END_VAR
VAR
    uiCh    : UINT;      // канал
    uiBits  : UINT;      // три бита канала
    xDemand : BOOL;      // требование канала
END_VAR

(* ---- RowInputs.method.impl.st ---- *)
// AUTO-GENERATED by cemgen 1.0.0 — не редактировать: правьте матрицу и запустите
//   python -m cemgen generate <файл матрицы .csv или .xlsx>
// Матрица: SIS-V101-CEM, объект V-101, ревизия B от 2026-10-19, SHA-256 сетки df2ed4841a9453ca
FOR uiCh := 1 TO GVL_Const.SIS_VOTE_CH_MAX DO
    uiBits := SEL(uiCh <= uiChannels, 0, SHR(uiRow, 3 * (uiCh - 1)) AND 7);
    xDemand := (uiBits AND 1) <> 0;
    stIn.axDi[uiCh] := NOT xDemand;
    stIn.axDiValid[uiCh] := (uiBits AND 2) <> 0;
    stIn.arAi_eu[uiCh] := SEL(xDemand, 40.0, 60.0);
    stIn.axAiValid[uiCh] := (uiBits AND 2) <> 0;
    stCmd.axBypassReq[uiCh] := xBypass AND ((uiBits AND 4) <> 0);
END_FOR

(* ---- RowStates.method.decl.st ---- *)
// AUTO-GENERATED by cemgen 1.0.0 — не редактировать: правьте матрицу и запустите
//   python -m cemgen generate <файл матрицы .csv или .xlsx>
// Матрица: SIS-V101-CEM, объект V-101, ревизия B от 2026-10-19, SHA-256 сетки df2ed4841a9453ca
// Назначение: вспомогательный метод набора FB_VoteTruth_Test.
// Автор:      kr0nsch; код — генератор cemgen
// Версия:     1.0.0
// Документ:   docs/DESIGN.md, раздел «10. Генератор cemgen»; docs/cause_effect_matrix.md
// ВНИМАНИЕ:   код демонстрационный и не предназначен для систем безопасности. Реальная ПАЗ требует
//             определения SIL, сертифицированных аппаратных и программных средств и валидации по
//             ГОСТ Р МЭК 61511.
// Состояния каналов строки уровня 1: код (r SHR 2(k − 1)) AND 3 — 0 Normal, 1 Demand, 2 Invalid, 3
// Bypassed; каналы k > N — NotUsed.
METHOD PRIVATE RowStates
VAR_INPUT
    uiRow      : UINT;   // строка таблицы
    uiChannels : UINT;   // N схемы
END_VAR
VAR_IN_OUT
    aeCh : ARRAY[1..GVL_Const.SIS_VOTE_CH_MAX] OF E_ChannelState;   // состояния каналов
END_VAR
VAR
    uiCh : UINT;         // канал
END_VAR

(* ---- RowStates.method.impl.st ---- *)
// AUTO-GENERATED by cemgen 1.0.0 — не редактировать: правьте матрицу и запустите
//   python -m cemgen generate <файл матрицы .csv или .xlsx>
// Матрица: SIS-V101-CEM, объект V-101, ревизия B от 2026-10-19, SHA-256 сетки df2ed4841a9453ca
FOR uiCh := 1 TO GVL_Const.SIS_VOTE_CH_MAX DO
    IF uiCh > uiChannels THEN
        aeCh[uiCh] := E_ChannelState.NotUsed;
    ELSE
        CASE SHR(uiRow, 2 * (uiCh - 1)) AND 3 OF
            0:
                aeCh[uiCh] := E_ChannelState.Normal;
            1:
                aeCh[uiCh] := E_ChannelState.Demand;
            2:
                aeCh[uiCh] := E_ChannelState.Invalid;
        ELSE
            aeCh[uiCh] := E_ChannelState.Bypassed;
        END_CASE
    END_IF
END_FOR
